(* IEC 61131-3 sources: llm-plc-st-eval/data/processed_definitivo/qwen2.5-coder_14b/B5/zero_shot, 3 files *)

(* ---- ejec_1.st ---- *)
FUNCTION_BLOCK FB_Ventilador
VAR_INPUT
    quemadorOn : BOOL; // Indica si el quemador está encendido
END_VAR

VAR_OUTPUT
    ventilador : BOOL; // Controla el ventilador
END_VAR

VAR
    timer : TON; // Timer de retardo
    timerDone : BOOL; // Indica si el timer ha terminado
END_VAR

// Inicialización del timer
IF NOT timerDone THEN
    timer(IN := NOT quemadorOn, PT := T#30S);
    timerDone := timer.Q;
END_IF;

// Control del ventilador
IF quemadorOn OR NOT timerDone THEN
    ventilador := TRUE;
ELSE
    ventilador := FALSE;
END_IF;

(* ---- ejec_2.st ---- *)
FUNCTION_BLOCK FB_Ventilador
VAR_INPUT
    quemadorOn : BOOL; // Estado del quemador (TRUE si encendido, FALSE si apagado)
END_VAR

VAR_OUTPUT
    ventilador : BOOL; // Estado del ventilador (TRUE si encendido, FALSE si apagado)
END_VAR

VAR
    timer : TON; // Timer de retardo
    timerDone : BOOL; // Bandera para indicar si el timer ha terminado
END_VAR

// Inicialización del timer
IF NOT timerDone THEN
    timer(IN := NOT quemadorOn, PT := T#30S);
    timerDone := timer.Q;
END_IF;

// Control del ventilador
IF quemadorOn OR (NOT quemadorOn AND NOT timerDone) THEN
    ventilador := TRUE;
ELSE
    ventilador := FALSE;
END_IF;

(* ---- ejec_3.st ---- *)
FUNCTION_BLOCK FB_Ventilador
VAR_INPUT
    quemadorOn : BOOL; // Estado del quemador (encendido/apagado)
END_VAR

VAR_OUTPUT
    ventilador : BOOL; // Estado del ventilador (encendido/apagado)
END_VAR

VAR
    timer : TON; // Timer de retardo
    timerDone : BOOL; // Bandera para indicar que el timer ha terminado
END_VAR

// Inicialización del timer
IF NOT timer.Q THEN
    timer(IN := FALSE, PT := T#30S);
END_IF;

// Lógica del ventilador
IF quemadorOn THEN
    ventilador := TRUE; // El ventilador se enciende cuando el quemador está encendido
    timer(IN := FALSE); // Reinicia el timer
ELSE
    IF NOT timer.Q THEN
        timer(IN := TRUE); // Inicia el timer cuando el quemador se apaga
    END_IF;
    ventilador := timer.Q; // El ventilador se apaga cuando el timer termina
END_IF;
